FUNCTION_BLOCK FB_Conveyor
VAR_OUTPUT
    motorRunning : BOOL;
    productCount : UDINT;
    alarm : STRING(80);
END_VAR
VAR
    requested : BOOL;
    configuredDelay : TIME := T#1s;
    startup : TON;
    productEdge : R_TRIG;
END_VAR


(* Invoke public methods explicitly. *)


METHOD PUBLIC Start
VAR_INPUT
    delay : TIME := T#1s;
END_VAR

configuredDelay := delay;
requested := TRUE;
END_METHOD


METHOD PUBLIC Stop

requested := FALSE;
startup(IN := FALSE, PT := configuredDelay);
motorRunning := FALSE;
alarm := 'Stopped';
END_METHOD


METHOD PUBLIC Reset

(* Reset the count while preserving the run command and sampled sensor edge. *)
productCount := 0;
END_METHOD


METHOD PUBLIC Update
VAR_INPUT
    guardClosed : BOOL;
    stopRequested : BOOL := FALSE;
    sensor : BOOL := FALSE;
END_VAR

(* Interlocks win even if Start was called earlier in this scan. *)
IF stopRequested OR NOT guardClosed THEN
    Stop();
END_IF;
startup(IN := requested, PT := configuredDelay);
motorRunning := startup.Q;
CountProduct(sensor := sensor);
IF NOT guardClosed THEN
    alarm := 'Guard open';
ELSIF stopRequested THEN
    alarm := 'Stopped';
ELSIF requested AND NOT motorRunning THEN
    alarm := 'Starting';
ELSE
    alarm := '';
END_IF;
END_METHOD


METHOD PUBLIC IsRunning : BOOL

IsRunning := motorRunning;
END_METHOD


METHOD PRIVATE CountProduct
VAR_INPUT
    sensor : BOOL;
END_VAR

(* Sampling also while stopped prevents a stale edge on restart. *)
productEdge(CLK := sensor);
IF motorRunning AND productEdge.Q THEN
    productCount := productCount + 1;
END_IF;
END_METHOD

END_FUNCTION_BLOCK

(* stored: Version 1.1.0.1, ProductVersion 3.1 *)
